Fanuc KAREL source: kt00585.KL

-- PROVISIONAL review KL for V940-1; original PC SHA256 2a1c3db6e27e56643cd3ac939a1ca8b51571fc00e5e21ae552e41e7d223a70e1
-- Incomplete behavior may be omitted. Consult companion uncertainty JSON. Do not deploy.
PROGRAM KT00585
%NOLOCKGROUP
VAR
  I1 : INTEGER
-- UNRESOLVED_DECL V2 type=000013
-- UNRESOLVED_DECL OUT type=000013
BEGIN
  -- V9_ZERO_TABLE_METADATA_HINT layout=0001; no indexed target words; source/name/runtime held
  -- UNRESOLVED_PC offsets 5-16; opcodes 2E,23
  -- UNRESOLVED_PC offsets 21-36; opcodes 2E,22,32,35
  -- UNRESOLVED_PC offsets 41-63; opcodes 21,49,8B,4A
  -- UNRESOLVED_PC offsets 68-72; opcodes 7F
END KT00585
